// TIA Portal V21 export
// export: Created 2026-11-10T19:11:38.7758442Z, ExportSetting WithDefaults, DisplayName Totally Integrated Automation Portal, DisplayVersion V21 Update 3, DisplayName STEP 7 Professional, DisplayVersion V21 Update 3, DisplayName STEP 7 Safety, DisplayVersion V21, DisplayName Tech WebApplication, DisplayVersion V21, DisplayName WinCC Basic/Comfort/Advanced, DisplayVersion V21 Update 3, DisplayName WinCC Unified, DisplayVersion V21 Update 3
DATA_BLOCK "DB_LEAD_LAG"   // DB27
// stored: AutoNumber true, DBAccessibleFromOPCUA true, DBAccessibleFromWebserver true, InstanceOfName LEAD_LAG, OfSystemLibElement LEAD_LAG, OfSystemLibVersion 2.1
"LEAD_LAG"
   // VAR_INPUT
   //    IN : Real;
   //    SAMPLE_T : Int;
   // END_VAR
   // VAR_OUTPUT
   //    OUT : Real;
   //    ERR_CODE : Word;
   // END_VAR
   // VAR
   //    LD_TIME : Real;
   //    GAIN : Real;
   //    PREV_IN : Real;
   //    PREV_OUT : Real;
   //    LG_TIME : Real;
   // END_VAR
BEGIN
END_DATA_BLOCK
